Staubli VAL3: getFrame.pgx

public program getFrame(num x_nIndex, frame& x_fFrame)
begin

  link(x_fFrame,world)
  x_fFrame=fFrameItem[x_nIndex].fFrame

end
